Yaskawa INFORM job: SIMPSTSQA.JBI

/JOB
//NAME SIMPSTSQA
//POS
///NPOS 227,0,0,0,0,0
///TOOL 0
///POSTYPE PULSE
///PULSE
C00000=181936,125599,48049,36468,-166396,-244514
C00001=91044,123269,-27074,-39529,-118967,-320932
C00002=91026,121985,-26720,-39399,-119901,-321366
C00003=91025,121902,-26696,-39391,-119962,-321395
C00004=84441,128980,-9878,-35943,-127586,-322187
C00005=84433,128997,-9839,-35939,-127603,-322190
C00006=84442,129005,-9823,-35941,-127607,-322195
C00007=84450,129013,-9807,-35945,-127612,-322202
C00008=131590,171329,90336,-11181,-176231,-305722
C00009=131604,171353,90383,-11188,-176249,-305732
C00010=131612,171347,90369,-11191,-176242,-305735
C00011=131620,171341,90355,-11195,-176236,-305740
C00012=130664,144233,24264,-32397,-141980,-324627
C00013=130676,144217,24227,-32402,-141964,-324627
C00014=130671,144206,24205,-32400,-141956,-324621
C00015=130666,144195,24183,-32398,-141949,-324616
C00016=98641,115570,-42335,-43643,-112674,-320477
C00017=98617,115560,-42354,-43634,-112671,-320468
C00018=98607,115565,-42342,-43628,-112677,-320468
C00019=98597,115569,-42330,-43623,-112684,-320468
C00020=91034,121894,-26715,-39395,-119953,-321394
C00021=91032,121811,-26692,-39387,-120014,-321423
C00022=84440,128902,-9856,-35938,-127644,-322212
C00023=84432,128920,-9816,-35934,-127661,-322215
C00024=84441,128927,-9801,-35937,-127665,-322220
C00025=84449,128935,-9785,-35940,-127670,-322224
C00026=116230,158955,57758,-26752,-157559,-322631
C00027=116247,158973,57792,-26759,-157569,-322642
C00028=116254,158966,57778,-26762,-157562,-322644
C00029=116262,158960,57764,-26765,-157555,-322647
C00030=130664,144164,24286,-32396,-142034,-324647
C00031=130676,144148,24249,-32401,-142017,-324647
C00032=130671,144137,24227,-32399,-142010,-324640
C00033=130666,144126,24205,-32397,-142002,-324635
C00034=98638,115482,-42310,-43630,-112738,-320511
C00035=98615,115472,-42328,-43621,-112735,-320502
C00036=98605,115477,-42316,-43615,-112741,-320502
C00037=98594,115481,-42304,-43610,-112747,-320502
C00038=91041,121803,-26711,-39391,-120005,-321421
C00039=84440,128892,-9853,-35938,-127652,-322215
C00040=84432,128910,-9814,-35933,-127668,-322218
C00041=84441,128917,-9798,-35936,-127673,-322223
C00042=84449,128925,-9782,-35939,-127677,-322228
C00043=116230,158931,57767,-26753,-157578,-322637
C00044=116247,158949,57801,-26760,-157588,-322649
C00045=116254,158943,57787,-26763,-157581,-322650
C00046=116262,158936,57772,-26766,-157574,-322652
C00047=130664,144121,24300,-32395,-142067,-324658
C00048=130676,144105,24263,-32401,-142051,-324658
C00049=130671,144094,24240,-32399,-142043,-324653
C00050=130666,144083,24218,-32397,-142036,-324648
C00051=98637,115405,-42287,-43619,-112794,-320541
C00052=98613,115395,-42306,-43609,-112791,-320531
C00053=98603,115400,-42294,-43604,-112797,-320531
C00054=98593,115404,-42281,-43599,-112803,-320531
C00055=91040,121720,-26687,-39383,-120066,-321449
C00056=84440,128815,-9830,-35933,-127710,-322237
C00057=84432,128832,-9791,-35928,-127726,-322242
C00058=84440,128840,-9775,-35931,-127731,-322247
C00059=84449,128847,-9759,-35934,-127736,-322252
C00060=116230,158869,57789,-26755,-157629,-322652
C00061=116247,158887,57824,-26762,-157639,-322663
C00062=116255,158880,57809,-26765,-157632,-322667
C00063=116262,158874,57795,-26768,-157625,-322668
C00064=130664,144052,24321,-32395,-142121,-324677
C00065=130676,144035,24284,-32400,-142104,-324677
C00066=130671,144025,24262,-32398,-142097,-324673
C00067=130666,144014,24240,-32396,-142089,-324668
C00068=98635,115317,-42261,-43606,-112858,-320575
C00069=98611,115307,-42280,-43597,-112854,-320565
C00070=98601,115312,-42268,-43591,-112861,-320565
C00071=98591,115316,-42256,-43586,-112867,-320565
C00072=91039,121637,-26663,-39375,-120127,-321478
C00073=84439,128737,-9808,-35928,-127768,-322262
C00074=84431,128754,-9768,-35923,-127785,-322265
C00075=84440,128762,-9752,-35926,-127789,-322271
C00076=84448,128770,-9737,-35929,-127794,-322276
C00077=116231,158807,57812,-26757,-157680,-322668
C00078=116247,158825,57847,-26764,-157690,-322679
C00079=116255,158818,57832,-26767,-157683,-322681
C00080=116263,158812,57818,-26770,-157676,-322683
C00081=130664,143983,24343,-32394,-142174,-324697
C00082=130676,143966,24306,-32399,-142158,-324697
C00083=130671,143956,24284,-32397,-142150,-324692
C00084=130666,143945,24262,-32395,-142143,-324687
C00085=98633,115229,-42235,-43593,-112921,-320609
C00086=98609,115219,-42254,-43584,-112918,-320599
C00087=98599,115224,-42242,-43578,-112924,-320599
C00088=98589,115228,-42230,-43573,-112931,-320599
C00089=91038,121554,-26639,-39367,-120188,-321506
C00090=84439,128659,-9785,-35923,-127826,-322286
C00091=84431,128676,-9746,-35918,-127843,-322289
C00092=84439,128684,-9730,-35921,-127847,-322294
C00093=84447,128692,-9714,-35924,-127852,-322301
C00094=116231,158744,57835,-26759,-157732,-322683
C00095=116247,158762,57870,-26766,-157742,-322694
C00096=116255,158756,57855,-26769,-157735,-322697
C00097=116263,158750,57841,-26772,-157728,-322699
C00098=130663,143914,24365,-32393,-142228,-324716
C00099=130676,143898,24328,-32398,-142211,-324716
C00100=130671,143887,24306,-32397,-142204,-324711
C00101=130666,143876,24284,-32395,-142196,-324707
C00102=98631,115141,-42209,-43580,-112985,-320643
C00103=98607,115131,-42228,-43571,-112982,-320633
C00104=98597,115136,-42216,-43566,-112988,-320633
C00105=98587,115140,-42203,-43561,-112994,-320633
C00106=91036,121471,-26615,-39358,-120249,-321535
C00107=84438,128581,-9762,-35918,-127885,-322310
C00108=84430,128598,-9723,-35913,-127901,-322314
C00109=84439,128606,-9707,-35917,-127906,-322318
C00110=84447,128614,-9691,-35919,-127910,-322325
C00111=116231,158682,57858,-26761,-157783,-322699
C00112=116247,158700,57893,-26768,-157793,-322710
C00113=116255,158694,57878,-26771,-157786,-322712
C00114=116263,158687,57864,-26774,-157779,-322713
C00115=130663,143845,24387,-32392,-142281,-324736
C00116=130676,143829,24350,-32398,-142265,-324736
C00117=130671,143818,24328,-32396,-142257,-324731
C00118=130666,143807,24306,-32394,-142250,-324726
C00119=98629,115053,-42183,-43567,-113049,-320677
C00120=98605,115043,-42202,-43558,-113046,-320667
C00121=98595,115048,-42190,-43553,-113052,-320665
C00122=98585,115053,-42177,-43548,-113058,-320665
C00123=91035,121389,-26590,-39350,-120310,-321562
C00124=84438,128503,-9739,-35913,-127943,-322335
C00125=84430,128521,-9700,-35909,-127959,-322338
C00126=84438,128529,-9684,-35912,-127964,-322343
C00127=84446,128536,-9668,-35915,-127969,-322348
C00128=116231,158620,57881,-26763,-157834,-322713
C00129=116247,158638,57916,-26770,-157844,-322725
C00130=116255,158632,57901,-26773,-157837,-322728
C00131=116263,158625,57887,-26776,-157830,-322730
C00132=130663,143776,24409,-32392,-142335,-324755
C00133=130676,143760,24373,-32397,-142319,-324755
C00134=130671,143749,24350,-32395,-142311,-324750
C00135=130666,143738,24328,-32393,-142304,-324745
C00136=98627,114965,-42157,-43555,-113113,-320711
C00137=98603,114956,-42176,-43546,-113110,-320699
C00138=98593,114960,-42163,-43540,-113116,-320699
C00139=98583,114965,-42151,-43535,-113122,-320699
C00140=91034,121306,-26566,-39342,-120371,-321591
C00141=84437,128426,-9716,-35908,-128001,-322357
C00142=84429,128443,-9677,-35904,-128018,-322362
C00143=84438,128451,-9661,-35907,-128022,-322367
C00144=84446,128459,-9645,-35910,-128027,-322372
C00145=116231,158558,57905,-26765,-157886,-322730
C00146=116247,158576,57939,-26772,-157896,-322741
C00147=116255,158570,57925,-26775,-157889,-322743
C00148=116263,158563,57910,-26778,-157882,-322746
C00149=130663,143707,24432,-32391,-142389,-324775
C00150=130676,143691,24395,-32396,-142372,-324775
C00151=130671,143680,24373,-32394,-142365,-324770
C00152=130666,143669,24350,-32392,-142357,-324765
C00153=98625,114878,-42130,-43542,-113177,-320745
C00154=98601,114868,-42149,-43533,-113173,-320733
C00155=98591,114872,-42137,-43528,-113180,-320733
C00156=98581,114877,-42125,-43522,-113186,-320733
C00157=91033,121224,-26542,-39334,-120433,-321619
C00158=84436,128348,-9693,-35904,-128060,-322382
C00159=84428,128366,-9654,-35899,-128076,-322385
C00160=84437,128374,-9638,-35902,-128081,-322391
C00161=84445,128381,-9622,-35905,-128085,-322396
C00162=116231,158496,57928,-26767,-157937,-322744
C00163=116248,158514,57963,-26774,-157947,-322757
C00164=116255,158508,57948,-26777,-157940,-322759
C00165=116263,158501,57934,-26780,-157933,-322760
C00166=130663,143638,24454,-32390,-142442,-324794
C00167=130676,143622,24417,-32395,-142426,-324794
C00168=130671,143611,24395,-32393,-142418,-324789
C00169=130666,143600,24373,-32391,-142411,-324784
C00170=98623,114790,-42104,-43530,-113240,-320777
C00171=98599,114780,-42123,-43520,-113237,-320767
C00172=98589,114785,-42111,-43515,-113244,-320767
C00173=98579,114789,-42099,-43510,-113250,-320767
C00174=91032,121141,-26517,-39326,-120494,-321648
C00175=84436,128271,-9670,-35899,-128118,-322406
C00176=84428,128288,-9630,-35894,-128135,-322409
C00177=84436,128296,-9614,-35897,-128139,-322416
C00178=84445,128304,-9599,-35900,-128144,-322420
C00179=116231,158434,57952,-26769,-157989,-322760
C00180=116248,158452,57986,-26776,-157999,-322772
C00181=116256,158446,57972,-26780,-157992,-322773
C00182=116263,158439,57957,-26782,-157985,-322777
C00183=130663,143570,24476,-32389,-142496,-324814
C00184=130676,143553,24440,-32395,-142480,-324814
C00185=130671,143543,24417,-32393,-142472,-324809
C00186=130666,143532,24395,-32391,-142465,-324804
C00187=98621,114702,-42077,-43517,-113304,-320811
C00188=98597,114692,-42096,-43508,-113301,-320801
C00189=98587,114697,-42084,-43502,-113308,-320801
C00190=98577,114702,-42072,-43497,-113314,-320801
C00191=91031,121058,-26492,-39318,-120555,-321676
C00192=84435,128193,-9646,-35894,-128177,-322430
C00193=84427,128211,-9607,-35889,-128193,-322433
C00194=84436,128219,-9591,-35892,-128198,-322438
C00195=84444,128226,-9575,-35895,-128202,-322445
C00196=116231,158372,57975,-26771,-158040,-322777
C00197=116248,158390,58010,-26779,-158050,-322788
C00198=116256,158384,57995,-26782,-158043,-322790
C00199=116264,158378,57981,-26785,-158036,-322791
C00200=130663,143501,24499,-32389,-142550,-324833
C00201=130676,143485,24462,-32394,-142533,-324833
C00202=130671,143474,24440,-32392,-142526,-324828
C00203=130666,143463,24418,-32390,-142518,-324823
C00204=98619,114615,-42051,-43504,-113368,-320845
C00205=98595,114605,-42070,-43495,-113365,-320835
C00206=98585,114610,-42057,-43490,-113372,-320835
C00207=98575,114614,-42045,-43485,-113378,-320835
C00208=91030,120976,-26468,-39309,-120616,-321703
C00209=84435,128116,-9623,-35889,-128235,-322454
C00210=84427,128133,-9584,-35885,-128252,-322458
C00211=84435,128141,-9568,-35888,-128256,-322463
C00212=84444,128149,-9552,-35891,-128261,-322469
C00213=116232,158310,57999,-26774,-158092,-322791
C00214=116248,158328,58034,-26781,-158102,-322803
C00215=116256,158322,58019,-26784,-158095,-322806
C00216=116264,158316,58005,-26787,-158088,-322807
C00217=130663,143432,24522,-32388,-142603,-324854
C00218=130676,143416,24485,-32393,-142587,-324854
C00219=130671,143405,24463,-32391,-142580,-324848
C00220=130666,143394,24440,-32389,-142572,-324843
C00221=98617,114527,-42024,-43492,-113432,-320879
C00222=98593,114517,-42043,-43483,-113429,-320869
C00223=98583,114522,-42031,-43477,-113436,-320869
C00224=98573,114527,-42019,-43472,-113442,-320869
C00225=91029,120894,-26443,-39301,-120677,-321732
C00226=107798,118362,10887,-23094,-151190,-316635
//INST
///DATE 2026/02/26 14:39
///COMM Generated using RoboDK
///ATTR SC,RW
///GROUP1 RB1
NOP
MOVJ C00000 VJ=50.00 PL=1
MOVL C00001 V=1000.0 PL=1
MOVL C00002 V=130.0 PL=1
MOVL C00003 V=130.0 PL=1
MOVL C00004 V=30.0 PL=1
MOVL C00005 V=30.0 PL=1
MOVL C00006 V=30.0 PL=1
MOVL C00007 V=30.0 PL=1
MOVL C00008 V=30.0 PL=1
MOVL C00009 V=30.0 PL=1
MOVL C00010 V=30.0 PL=1
MOVL C00011 V=30.0 PL=1
MOVL C00012 V=30.0 PL=1
MOVL C00013 V=30.0 PL=1
MOVL C00014 V=30.0 PL=1
MOVL C00015 V=30.0 PL=1
MOVL C00016 V=30.0 PL=1
MOVL C00017 V=30.0 PL=1
MOVL C00018 V=30.0 PL=1
MOVL C00019 V=30.0 PL=1
MOVL C00020 V=30.0 PL=1
MOVL C00021 V=130.0 PL=1
MOVL C00022 V=30.0 PL=1
MOVL C00023 V=30.0 PL=1
MOVL C00024 V=30.0 PL=1
MOVL C00025 V=30.0 PL=1
MOVL C00026 V=30.0 PL=1
MOVL C00027 V=30.0 PL=1
MOVL C00028 V=30.0 PL=1
MOVL C00029 V=30.0 PL=1
MOVL C00030 V=30.0 PL=1
MOVL C00031 V=30.0 PL=1
MOVL C00032 V=30.0 PL=1
MOVL C00033 V=30.0 PL=1
MOVL C00034 V=30.0 PL=1
MOVL C00035 V=30.0 PL=1
MOVL C00036 V=30.0 PL=1
MOVL C00037 V=30.0 PL=1
MOVL C00038 V=30.0 PL=1
MOVL C00039 V=30.0 PL=1
MOVL C00040 V=30.0 PL=1
MOVL C00041 V=30.0 PL=1
MOVL C00042 V=30.0 PL=1
MOVL C00043 V=30.0 PL=1
MOVL C00044 V=30.0 PL=1
MOVL C00045 V=30.0 PL=1
MOVL C00046 V=30.0 PL=1
MOVL C00047 V=30.0 PL=1
MOVL C00048 V=30.0 PL=1
MOVL C00049 V=30.0 PL=1
MOVL C00050 V=30.0 PL=1
MOVL C00051 V=30.0 PL=1
MOVL C00052 V=30.0 PL=1
MOVL C00053 V=30.0 PL=1
MOVL C00054 V=30.0 PL=1
MOVL C00055 V=30.0 PL=1
MOVL C00056 V=30.0 PL=1
MOVL C00057 V=30.0 PL=1
MOVL C00058 V=30.0 PL=1
MOVL C00059 V=30.0 PL=1
MOVL C00060 V=30.0 PL=1
MOVL C00061 V=30.0 PL=1
MOVL C00062 V=30.0 PL=1
MOVL C00063 V=30.0 PL=1
MOVL C00064 V=30.0 PL=1
MOVL C00065 V=30.0 PL=1
MOVL C00066 V=30.0 PL=1
MOVL C00067 V=30.0 PL=1
MOVL C00068 V=30.0 PL=1
MOVL C00069 V=30.0 PL=1
MOVL C00070 V=30.0 PL=1
MOVL C00071 V=30.0 PL=1
MOVL C00072 V=30.0 PL=1
MOVL C00073 V=30.0 PL=1
MOVL C00074 V=30.0 PL=1
MOVL C00075 V=30.0 PL=1
MOVL C00076 V=30.0 PL=1
MOVL C00077 V=30.0 PL=1
MOVL C00078 V=30.0 PL=1
MOVL C00079 V=30.0 PL=1
MOVL C00080 V=30.0 PL=1
MOVL C00081 V=30.0 PL=1
MOVL C00082 V=30.0 PL=1
MOVL C00083 V=30.0 PL=1
MOVL C00084 V=30.0 PL=1
MOVL C00085 V=30.0 PL=1
MOVL C00086 V=30.0 PL=1
MOVL C00087 V=30.0 PL=1
MOVL C00088 V=30.0 PL=1
MOVL C00089 V=30.0 PL=1
MOVL C00090 V=30.0 PL=1
MOVL C00091 V=30.0 PL=1
MOVL C00092 V=30.0 PL=1
MOVL C00093 V=30.0 PL=1
MOVL C00094 V=30.0 PL=1
MOVL C00095 V=30.0 PL=1
MOVL C00096 V=30.0 PL=1
MOVL C00097 V=30.0 PL=1
MOVL C00098 V=30.0 PL=1
MOVL C00099 V=30.0 PL=1
MOVL C00100 V=30.0 PL=1
MOVL C00101 V=30.0 PL=1
MOVL C00102 V=30.0 PL=1
MOVL C00103 V=30.0 PL=1
MOVL C00104 V=30.0 PL=1
MOVL C00105 V=30.0 PL=1
MOVL C00106 V=30.0 PL=1
MOVL C00107 V=30.0 PL=1
MOVL C00108 V=30.0 PL=1
MOVL C00109 V=30.0 PL=1
MOVL C00110 V=30.0 PL=1
MOVL C00111 V=30.0 PL=1
MOVL C00112 V=30.0 PL=1
MOVL C00113 V=30.0 PL=1
MOVL C00114 V=30.0 PL=1
MOVL C00115 V=30.0 PL=1
MOVL C00116 V=30.0 PL=1
MOVL C00117 V=30.0 PL=1
MOVL C00118 V=30.0 PL=1
MOVL C00119 V=30.0 PL=1
MOVL C00120 V=30.0 PL=1
MOVL C00121 V=30.0 PL=1
MOVL C00122 V=30.0 PL=1
MOVL C00123 V=30.0 PL=1
MOVL C00124 V=30.0 PL=1
MOVL C00125 V=30.0 PL=1
MOVL C00126 V=30.0 PL=1
MOVL C00127 V=30.0 PL=1
MOVL C00128 V=30.0 PL=1
MOVL C00129 V=30.0 PL=1
MOVL C00130 V=30.0 PL=1
MOVL C00131 V=30.0 PL=1
MOVL C00132 V=30.0 PL=1
MOVL C00133 V=30.0 PL=1
MOVL C00134 V=30.0 PL=1
MOVL C00135 V=30.0 PL=1
MOVL C00136 V=30.0 PL=1
MOVL C00137 V=30.0 PL=1
MOVL C00138 V=30.0 PL=1
MOVL C00139 V=30.0 PL=1
MOVL C00140 V=30.0 PL=1
MOVL C00141 V=30.0 PL=1
MOVL C00142 V=30.0 PL=1
MOVL C00143 V=30.0 PL=1
MOVL C00144 V=30.0 PL=1
MOVL C00145 V=30.0 PL=1
MOVL C00146 V=30.0 PL=1
MOVL C00147 V=30.0 PL=1
MOVL C00148 V=30.0 PL=1
MOVL C00149 V=30.0 PL=1
MOVL C00150 V=30.0 PL=1
MOVL C00151 V=30.0 PL=1
MOVL C00152 V=30.0 PL=1
MOVL C00153 V=30.0 PL=1
MOVL C00154 V=30.0 PL=1
MOVL C00155 V=30.0 PL=1
MOVL C00156 V=30.0 PL=1
MOVL C00157 V=30.0 PL=1
MOVL C00158 V=30.0 PL=1
MOVL C00159 V=30.0 PL=1
MOVL C00160 V=30.0 PL=1
MOVL C00161 V=30.0 PL=1
MOVL C00162 V=30.0 PL=1
MOVL C00163 V=30.0 PL=1
MOVL C00164 V=30.0 PL=1
MOVL C00165 V=30.0 PL=1
MOVL C00166 V=30.0 PL=1
MOVL C00167 V=30.0 PL=1
MOVL C00168 V=30.0 PL=1
MOVL C00169 V=30.0 PL=1
MOVL C00170 V=30.0 PL=1
MOVL C00171 V=30.0 PL=1
MOVL C00172 V=30.0 PL=1
MOVL C00173 V=30.0 PL=1
MOVL C00174 V=30.0 PL=1
MOVL C00175 V=30.0 PL=1
MOVL C00176 V=30.0 PL=1
MOVL C00177 V=30.0 PL=1
MOVL C00178 V=30.0 PL=1
MOVL C00179 V=30.0 PL=1
MOVL C00180 V=30.0 PL=1
MOVL C00181 V=30.0 PL=1
MOVL C00182 V=30.0 PL=1
MOVL C00183 V=30.0 PL=1
MOVL C00184 V=30.0 PL=1
MOVL C00185 V=30.0 PL=1
MOVL C00186 V=30.0 PL=1
MOVL C00187 V=30.0 PL=1
MOVL C00188 V=30.0 PL=1
MOVL C00189 V=30.0 PL=1
MOVL C00190 V=30.0 PL=1
MOVL C00191 V=30.0 PL=1
MOVL C00192 V=30.0 PL=1
MOVL C00193 V=30.0 PL=1
MOVL C00194 V=30.0 PL=1
MOVL C00195 V=30.0 PL=1
MOVL C00196 V=30.0 PL=1
MOVL C00197 V=30.0 PL=1
MOVL C00198 V=30.0 PL=1
MOVL C00199 V=30.0 PL=1
MOVL C00200 V=30.0 PL=1
MOVL C00201 V=30.0 PL=1
MOVL C00202 V=30.0 PL=1
MOVL C00203 V=30.0 PL=1
MOVL C00204 V=30.0 PL=1
MOVL C00205 V=30.0 PL=1
MOVL C00206 V=30.0 PL=1
MOVL C00207 V=30.0 PL=1
MOVL C00208 V=30.0 PL=1
MOVL C00209 V=30.0 PL=1
MOVL C00210 V=30.0 PL=1
MOVL C00211 V=30.0 PL=1
MOVL C00212 V=30.0 PL=1
MOVL C00213 V=30.0 PL=1
MOVL C00214 V=30.0 PL=1
MOVL C00215 V=30.0 PL=1
MOVL C00216 V=30.0 PL=1
MOVL C00217 V=30.0 PL=1
MOVL C00218 V=30.0 PL=1
MOVL C00219 V=30.0 PL=1
MOVL C00220 V=30.0 PL=1
MOVL C00221 V=30.0 PL=1
MOVL C00222 V=30.0 PL=1
MOVL C00223 V=30.0 PL=1
MOVL C00224 V=30.0 PL=1
MOVL C00225 V=30.0 PL=1
MOVL C00226 V=1000.0 PL=1
END
